(* IEC 61131-3 sources: kns-port-domestic/tools/plcopen/tests/fixtures/constructs/src/POUs/Devices/FB_Valve, 5 files *)

(* ---- FB_Valve.decl.st ---- *)
// Назначение: задвижка — FINAL-наследник базы с двумя интерфейсами
// Автор:      <ИМЯ ФАМИЛИЯ>
// Версия:     0.1.0
// Документ:   docs/plcopen.md
FUNCTION_BLOCK FINAL FB_Valve EXTENDS FB_DeviceBase IMPLEMENTS I_Positioner, I_Lockable
VAR_OUTPUT
    rPos_pct : REAL;
    xLocked : BOOL;
END_VAR
VAR
    rSetpoint_pct : REAL;
END_VAR
VAR CONSTANT
    POS_MAX : REAL := 100.0;
END_VAR

(* ---- FB_Valve.impl.st ---- *)
SUPER^();
IF NOT xLocked THEN
    rPos_pct := F_Clamp(rValue := rSetpoint_pct, rMin := 0.0, rMax := POS_MAX);
END_IF

(* ---- Lock.method.decl.st ---- *)
METHOD PUBLIC Lock
VAR_INPUT
    xLock : BOOL;
END_VAR

(* ---- MoveTo.method.decl.st ---- *)
METHOD PUBLIC MoveTo : BOOL
VAR_INPUT
    rPos_pct : REAL;
END_VAR
VAR_OUTPUT
    xDone : BOOL;
END_VAR

(* ---- Trace.method.decl.st ---- *)
// Внутренний метод библиотеки
METHOD INTERNAL Trace : ST_MotorCmd
VAR_IN_OUT
    stLast : ST_MotorCmd;
END_VAR
